Fanuc KAREL source: KT00111.KL

PROGRAM KT00111
%NOLOCKGROUP
VAR
  R1: REAL
  H2: ARRAY[2] OF SHORT
  OUT: INTEGER
BEGIN
  R1 = 2.0
    H2[1] = 3
  OUT = R1 / H2[1]
END KT00111
